// TIA Portal V19 export
// export: Created 2026-10-15T09:44:24.8579522Z, ExportSetting WithDefaults, DisplayName Totally Integrated Automation Portal, DisplayVersion V19, DisplayName TIA Portal Openness, DisplayVersion V19, DisplayName TIA Portal Version Control Interface, DisplayVersion V19, DisplayName STEP 7 Professional, DisplayVersion V19, DisplayName STEP 7 Safety, DisplayVersion V19, DisplayName WinCC Basic/Comfort/Advanced, DisplayVersion V19, DisplayName WinCC Unified, DisplayVersion V19
FUNCTION "ROLL_PB23" : Void   // FC30, SCL
{ S7_Optimized_Access := 'TRUE' }
VERSION : 0.1
// stored: AutoNumber true, IsIECCheckEnabled false, SetENOAutomatically false, UDAEnableTagReadback false
   VAR_TEMP
      r : Bool;
      a1 : Word;
      a2 : Word;
      activeDataBlock : Int;
      comparisonResults : Array[0..0] of Bool;
   END_VAR
BEGIN

   #r := FALSE;
   #a1 := W#16#0000;
   #a2 := W#16#0000;
   #activeDataBlock := 0;
   // PB23, STEP 5 network 1
   #activeDataBlock := 15;
   // PB23, STEP 5 network 2
   #r := (("ROLL_State".M[40, 3] OR "ROLL_State".M[40, 4] OR "ROLL_State".M[40, 5]) AND "ROLL_State".M[111, 4]);
   "ROLL_State".M[240, 0] := #r;
   // PB23, STEP 5 network 3
   #a2 := #a1;
   #a1 := W#16#2120;
   #r := "ROLL_State".M[240, 0];
   "ROLL_TimerOp"(Number := 51,
                  Operation := 1,
                  Signal := #r,
                  Preset := #a1);
   #r := "ROLL_State".S5Timers[51].Q;
   "ROLL_IO".Output[19, 0] := #r;
   // PB23, STEP 5 network 4
   #a2 := #a1;
   #a1 := W#16#1050;
   #r := ((NOT "ROLL_State".M[6, 1]) AND ("ROLL_State".M[40, 4] OR "ROLL_State".M[40, 5]) AND "ROLL_IO".Output[19, 0] AND "ROLL_State".M[240, 0] AND "ROLL_State".M[35, 2] AND "ROLL_State".S5Timers[70].Q);
   "ROLL_TimerOp"(Number := 52,
                  Operation := 0,
                  Signal := #r,
                  Preset := #a1);
   #r := "ROLL_State".S5Timers[52].Q;
   "ROLL_IO".Output[19, 1] := #r;
   // PB23, STEP 5 network 5
   #r := ("ROLL_IO".Input[0, 2] AND "ROLL_IO".Input[0, 4]);
   IF #r THEN
       "ROLL_State".M[103, 7] := TRUE;
   END_IF;
   #r := (NOT "ROLL_State".S5Timers[59].Q);
   IF #r THEN
       "ROLL_State".M[103, 7] := FALSE;
   END_IF;
   // PB23, STEP 5 network 6
   #a2 := #a1;
   #a1 := W#16#3360;
   #r := "ROLL_State".S5Timers[59].Q;
   "ROLL_TimerOp"(Number := 76,
                  Operation := 0,
                  Signal := #r,
                  Preset := #a1);
   // PB23, STEP 5 network 7
   #r := ((NOT "ROLL_State".M[13, 3]) AND (NOT "ROLL_State".M[5, 6]) AND (NOT "ROLL_State".M[6, 2]) AND (NOT "ROLL_State".M[6, 3]) AND (((NOT "ROLL_State".S5Timers[76].Q) AND "ROLL_IO".Input[2, 2]) OR "ROLL_State".M[103, 7] OR "ROLL_State".M[152, 0]) AND ("ROLL_IO".Input[2, 2] OR "ROLL_State".M[152, 0]) AND "ROLL_IO".Input[3, 4] AND "ROLL_IO".Input[5, 6] AND "ROLL_State".S5Timers[59].Q);
   "ROLL_IO".Output[19, 5] := #r;
   // PB23, STEP 5 network 8
   #r := ((NOT "ROLL_State".M[5, 6]) AND (NOT "ROLL_State".M[6, 1]) AND ("ROLL_IO".Input[0, 1] OR "ROLL_IO".Input[0, 2]) AND "ROLL_IO".Input[3, 1] AND "ROLL_IO".Input[3, 4] AND "ROLL_State".M[0, 3] AND "ROLL_State".M[100, 0] AND "ROLL_State".S5Timers[70].Q);
   "ROLL_State".M[240, 0] := #r;
   // PB23, STEP 5 network 9
   #r := ((NOT "ROLL_IO".Output[20, 6]) AND (NOT "ROLL_State".M[5, 6]) AND (NOT "ROLL_State".M[8, 5]) AND (NOT "ROLL_State".S5Timers[96].Q) AND (("ROLL_State".M[100, 0] AND "ROLL_State".M[103, 1]) OR "ROLL_State".M[102, 6] OR "ROLL_State".M[104, 6]));
   "ROLL_IO".Output[20, 4] := #r;
   "ROLL_IO".Output[22, 6] := #r;
   // PB23, STEP 5 network 10
   #r := ((NOT "ROLL_IO".Output[20, 1]) AND ("ROLL_State".M[104, 0] OR "ROLL_State".M[104, 1] OR "ROLL_State".M[104, 4] OR "ROLL_State".M[152, 1]) AND "ROLL_State".M[99, 7]);
   "ROLL_IO".Output[20, 6] := #r;
   // PB23, STEP 5 network 11
   #r := ("ROLL_State".M[102, 7] OR "ROLL_State".M[103, 2] OR "ROLL_State".M[104, 5]);
   "ROLL_State".M[240, 0] := #r;
   // PB23, STEP 5 network 12
   #r := ((NOT "ROLL_State".M[13, 4]) AND (NOT "ROLL_State".M[6, 0]) AND (NOT "ROLL_State".M[6, 2]) AND (NOT "ROLL_State".M[7, 7]) AND "ROLL_IO".Input[3, 1] AND "ROLL_IO".Input[5, 0] AND "ROLL_IO".Input[5, 2] AND "ROLL_IO".Input[5, 4] AND "ROLL_State".M[240, 0]);
   "ROLL_IO".Output[20, 1] := #r;
   // PB23, STEP 5 network 13
   #r := "ROLL_State".M[103, 1];
   "ROLL_IO".Output[22, 2] := #r;
   // PB23, STEP 5 network 14
   #r := ("ROLL_State".M[102, 1] OR "ROLL_State".M[102, 2] OR "ROLL_State".M[102, 3] OR "ROLL_State".M[102, 6] OR "ROLL_State".M[102, 7] OR "ROLL_State".M[103, 2]);
   "ROLL_IO".Output[22, 3] := #r;
   // PB23, STEP 5 network 15
   #r := "ROLL_State".S5Timers[85].Q;
   "ROLL_IO".Output[21, 3] := #r;
   // PB23, STEP 5 network 16
   #a2 := #a1;
   #a1 := W#16#1020;
   #r := "ROLL_IO".Output[20, 6];
   "ROLL_TimerOp"(Number := 47,
                  Operation := 1,
                  Signal := #r,
                  Preset := #a1);
   // PB23, STEP 5 network 17
   #r := ((NOT "ROLL_IO".Output[21, 5]) AND (NOT "ROLL_IO".Output[22, 3]) AND (NOT "ROLL_IO".Output[22, 6]) AND (("ROLL_IO".Output[21, 4] AND "ROLL_State".S5Timers[47].Q) OR "ROLL_State".M[104, 0] OR "ROLL_State".M[152, 1]));
   "ROLL_IO".Output[21, 4] := #r;
   // PB23, STEP 5 network 18
   #r := ((NOT "ROLL_IO".Output[21, 4]) AND "ROLL_State".M[152, 0]);
   "ROLL_IO".Output[21, 5] := #r;
   // PB23, STEP 5 network 19
   RETURN;
END_FUNCTION
